FUNCTION_BLOCK FB_DeltaTime
(*
	Time since this instance was last called, in seconds. Call once per scan.
	Used by filters, ramps and controllers so they work at any task cycle time.
	Returns 0 on the first call.
*)
VAR_OUTPUT
	seconds					: LREAL; //seconds since the previous call
END_VAR
VAR
	lastTime			: ULINT; //system time of the previous call (100 ns units)
END_VAR

Update();

METHOD PROTECTED Update
VAR
	now : ULINT; //current system time (100 ns units)
END_VAR
now := F_GetSystemTime();
IF lastTime = 0 OR now < lastTime THEN
	seconds := 0;
ELSE
	seconds := ULINT_TO_LREAL(now - lastTime) * 1E-7;
END_IF
lastTime := now;
END_METHOD

END_FUNCTION_BLOCK

(* stored: Version 1.1.0.1, ProductVersion 3.1.4024.12
   POU FB_DeltaTime: Id {13b6bf83-6c01-4540-b1bd-4c7d86ecca35}, SpecialFunc None
   Folder Protected: Id {b7158dc9-66ef-4a5f-93ba-7395cdd4af00}
   Folder Logic: Id {b503138e-017b-4bca-8c54-22d85192c217}
   Method Update: Id {e236c7ba-3c0c-41f9-9a07-fbe7af51ff44} *)
